FUNCTION_BLOCK FsMove (* Rename, move or copy a file or directory on the file server *)
  (* Standard: 61499-2; Description: Uses iso_FscMoveFile() of the CCI ISOBUS driver (ISO 11783-13). The server copies or moves itself, no data goes over the bus. \n Client is NmDestin.s16OwnCfHnd, file server is NmDestin.s16Handle (e.g. found with NmGetCfInfo, NAME function 61). \n The FB opens its own io channel to the server and closes it at the end. One job at a time: REQ during a job gives ERR with s16Status E_BUSY. \n Every REQ ends with exactly one CNF or ERR. *)
  (* Version 1.0, 2026-11-26, Franz Höpfinger, initial API and implementation and/or initial documentation *)
  PACKAGE isobus::fs;
  IMPORT isobus::pgn::ISONETEVENT_T;
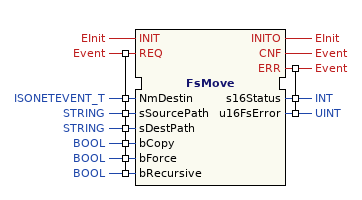
  EVENT_INPUT
    INIT : EInit; (* Service Initialization *)
    REQ WITH NmDestin, sSourcePath, sDestPath, bCopy, bForce, bRecursive; (* Move or copy *)
  END_EVENT
  EVENT_OUTPUT
    INITO : EInit; (* Initialization Confirm *)
    CNF; (* Moved or copied *)
    ERR WITH s16Status, u16FsError; (* Job failed *)
  END_EVENT
  VAR_INPUT
    NmDestin : isobus::pgn::ISONETEVENT_T; (* Client (s16OwnCfHnd) and file server (s16Handle) *)
    sSourcePath : STRING; (* Source on the file server *)
    sDestPath : STRING; (* Destination on the file server *)
    bCopy : BOOL; (* TRUE: copy instead of move *)
    bForce : BOOL; (* TRUE: overwrite an existing destination *)
    bRecursive : BOOL; (* TRUE: directory with its content *)
  END_VAR
  VAR_OUTPUT
    s16Status : INT; (* With ERR: driver return value or own error (E_BUSY, E_RANGE, E_CONFIG) *)
    u16FsError : UINT; (* With ERR: file server or client error (ISO 11783-13 B.9, 6400 ff. client) *)
  END_VAR
END_FUNCTION_BLOCK
